Fanuc KAREL source: KT00485.KL

PROGRAM KT00485
%NOLOCKGROUP
VAR
  P1: POSITION
  P2: XYZWPREXT
  OUT: XYZWPR
BEGIN
    P2.Y = 2.0
  OUT = P1 : P2
END KT00485
